{attribute 'call_after_init'}
FUNCTION_BLOCK FB_Conveyor EXTENDS FB_ConveyorBase
VAR_OUTPUT
    derivedInitCount : DINT;
END_VAR

SUPER^();

METHOD PUBLIC FB_init : BOOL
VAR_INPUT
    bInitRetains : BOOL;
    bInCopyCode : BOOL;
    conveyorId : DINT;
    sharedConfig : REFERENCE TO ST_ConveyorConfig;
    defaultDelay : TIME := T#100ms;
END_VAR
StartDelay := defaultDelay;
derivedInitCount := derivedInitCount + 1;
initTrace := initTrace * 10 + 2;
FB_init := TRUE;
END_METHOD

{attribute 'call_after_init'}
METHOD PUBLIC AfterInit
SUPER^.AfterInit();
initTrace := initTrace * 10 + 5;
ready := __ISVALIDREF(config) AND_THEN (id > 0 AND StartDelay > T#0ms AND factor > 0.0);
END_METHOD

END_FUNCTION_BLOCK

(* stored: Version 1.1.0.1, ProductVersion 3.1 *)
